(* IEC 61131-3 sources: tsplc/packages/build/tests/fixtures/raw-st/src/filling, 2 files *)

(* ---- E_StationState.st ---- *)
{attribute 'qualified_only'}
{attribute 'strict'}
TYPE E_StationState : (Idle := 0, Working := 1) USINT;
END_TYPE

(* ---- ST_Job.st ---- *)
TYPE ST_Job :
STRUCT
	Id : UDINT;
	Measurements : ARRAY [1..4] OF REAL;
END_STRUCT
END_TYPE
